(* PLC project Vn_nest_not, Beckhoff Automation GmbH TwinCAT PLC Control 3.5.13.21 *)
(* stored: creationDateTime 1970-01-01T00:00:00 *)

PROGRAM Vn_nest_not

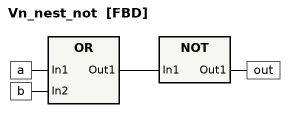
(* FBD diagram, written out as Structured Text *)
out := NOT (a OR b);
END_PROGRAM
